SUBAPPLICATION Uebung_OPC_L06_AX (* Wie Training_06 (Adapter-Variante von 04), lokal: Set/Reset/Toggle per localhost, Zustand lokal per PUBLISH *)
  (* Standard: 61499-2; Description: Copyright (c) 2026 Meisterschulen am Ostbahnhof This program and the accompanying materials are made available under the terms of the Eclipse Public License 2.0 which is available at https://www.eclipse.org/legal/epl-2.0/ SPDX-License-Identifier: EPL-2.0 *)
  (* Version 1.0, 2026-10-18, Franz Höpfinger, Meisterschulen am Ostbahnhof, Aus SubApp_PC_A + SubApp_PC_B von test_VV zusammengefuehrt, lokale Varianten der Bausteine *)
  PACKAGE Meins::OPC_UA_Lokal;
  IMPORT Uebungen::const::UT::DefaultPool::SoftKey_F1;
  IMPORT Uebungen::const::UT::DefaultPool::SoftKey_F2;
  IMPORT Uebungen::const::UT::DefaultPool::SoftKey_F3;
  IMPORT Meins::OPC_UA_Lokal::const::OpcUaLokal::SR1_SET_CALL;
  IMPORT Meins::OPC_UA_Lokal::const::OpcUaLokal::SR1_RESET_CALL;
  IMPORT Meins::OPC_UA_Lokal::const::OpcUaLokal::SR1_TOGGLE_CALL;
  IMPORT Meins::OPC_UA_Lokal::const::OpcUaLokal::SR1_STATE_READ;
  IMPORT logiBUS::io::DQ::logiBUS_DO::Output_Q1;
  IMPORT Meins::OPC_UA_Lokal::const::OpcUaLokal::SR1_SET_METHOD;
  IMPORT Meins::OPC_UA_Lokal::const::OpcUaLokal::SR1_RESET_METHOD;
  IMPORT Meins::OPC_UA_Lokal::const::OpcUaLokal::SR1_TOGGLE_METHOD;
  IMPORT Meins::OPC_UA_Lokal::const::OpcUaLokal::SR1_STATE_WRITE;
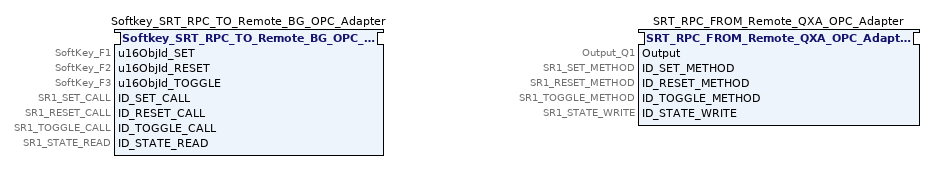
  SUBAPPS
    Softkey_SRT_RPC_TO_Remote_BG_OPC_Adapter : MyLib::sys::Softkey_SRT_RPC_TO_Remote_BG_OPC_Adapter(u16ObjId_SET := SoftKey_F1, u16ObjId_RESET := SoftKey_F2, u16ObjId_TOGGLE := SoftKey_F3, ID_SET_CALL := SR1_SET_CALL, ID_RESET_CALL := SR1_RESET_CALL, ID_TOGGLE_CALL := SR1_TOGGLE_CALL, ID_STATE_READ := SR1_STATE_READ);
    SRT_RPC_FROM_Remote_QXA_OPC_Adapter : MyLib::sys::SRT_RPC_FROM_Remote_QXA_OPC_Adapter_LOC(Output := Output_Q1, ID_SET_METHOD := SR1_SET_METHOD, ID_RESET_METHOD := SR1_RESET_METHOD, ID_TOGGLE_METHOD := SR1_TOGGLE_METHOD, ID_STATE_WRITE := SR1_STATE_WRITE);
  END_SUBAPPS
END_SUBAPPLICATION
